// TIA Portal V19 export
FUNCTION_BLOCK "RUA_R4"   // FB22, LAD
{ S7_Optimized_Access := 'TRUE' }
// stored: MemoryReserve 100, SetENOAutomatically false
   VAR
      START_Instance { S7_SetPoint := 'True'} : "START";
      "HEAT/COOL_Instance" { S7_SetPoint := 'True'} : "HEAT/COOL";
      "AUTO_COOLING_UTIITY SELECTION_Instance" { S7_SetPoint := 'True'} : "AUTO_COOLING_UTIITY SELECTION";
      AUTO_HEATING_SELECTION_Instance { S7_SetPoint := 'True'} : "AUTO_HEATING_SELECTION";
      "SEMI/_AUTO_Instance" { S7_SetPoint := 'True'} : "SEMI/_AUTO";
      COOLING_PROCESS_Instance { S7_SetPoint := 'True'} : "COOLING_PROCESS";
      HEATING_PROCEES_Instance { S7_SetPoint := 'True'} : "HEATING_PROCEES";
      RAMP_Instance { S7_SetPoint := 'True'} : "RAMP";
   END_VAR
BEGIN

REGION Network 1: START
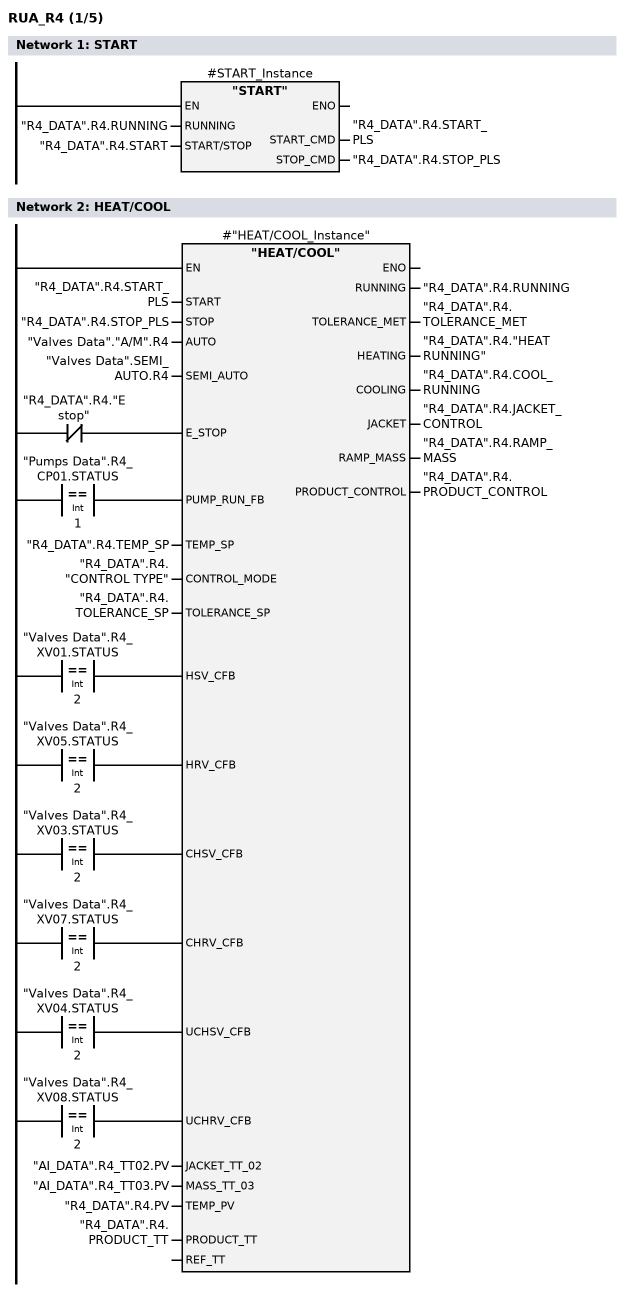
   RUNG wire#powerrail
      #START_Instance(RUNNING := "R4_DATA".R4.RUNNING, "START/STOP" := "R4_DATA".R4.START, START_CMD => "R4_DATA".R4.START_PLS, STOP_CMD => "R4_DATA".R4.STOP_PLS)
   END_RUNG
   // the same network as SCL:
   #START_Instance(RUNNING := "R4_DATA".R4.RUNNING,   // "START"
                   "START/STOP" := "R4_DATA".R4.START,
                   START_CMD => "R4_DATA".R4.START_PLS,
                   STOP_CMD => "R4_DATA".R4.STOP_PLS);
END_REGION

REGION Network 2: HEAT/COOL
   RUNG wire#powerrail
      #"HEAT/COOL_Instance"(E_STOP := wire#w1, PUMP_RUN_FB := wire#w2, HSV_CFB := wire#w3, HRV_CFB := wire#w4, CHSV_CFB := wire#w5, CHRV_CFB := wire#w6, UCHSV_CFB := wire#w7, UCHRV_CFB := wire#w8, START := "R4_DATA".R4.START_PLS, STOP := "R4_DATA".R4.STOP_PLS, AUTO := "Valves Data"."A/M".R4, SEMI_AUTO := "Valves Data".SEMI_AUTO.R4, TEMP_SP := "R4_DATA".R4.TEMP_SP, CONTROL_MODE := "R4_DATA".R4."CONTROL TYPE", TOLERANCE_SP := "R4_DATA".R4.TOLERANCE_SP, JACKET_TT_02 := "AI_DATA".R4_TT02.PV, MASS_TT_03 := "AI_DATA".R4_TT03.PV, TEMP_PV := "R4_DATA".R4.PV, PRODUCT_TT := "R4_DATA".R4.PRODUCT_TT, REF_TT :=, RUNNING => "R4_DATA".R4.RUNNING, TOLERANCE_MET => "R4_DATA".R4.TOLERANCE_MET, HEATING => "R4_DATA".R4."HEAT RUNNING", COOLING => "R4_DATA".R4.COOL_RUNNING, JACKET => "R4_DATA".R4.JACKET_CONTROL, RAMP_MASS => "R4_DATA".R4.RAMP_MASS, PRODUCT_CONTROL => "R4_DATA".R4.PRODUCT_CONTROL)
   END_RUNG
   RUNG wire#powerrail
      I_Contact( "R4_DATA".R4."E stop" )
   END_RUNG wire#w1
   RUNG wire#powerrail
      { S7_Templates := "SrcType := Int" } EQ_Contact(in1 := "Pumps Data".R4_CP01.STATUS, in2 := 1)
   END_RUNG wire#w2
   RUNG wire#powerrail
      { S7_Templates := "SrcType := Int" } EQ_Contact(in1 := "Valves Data".R4_XV01.STATUS, in2 := 2)
   END_RUNG wire#w3
   RUNG wire#powerrail
      { S7_Templates := "SrcType := Int" } EQ_Contact(in1 := "Valves Data".R4_XV05.STATUS, in2 := 2)
   END_RUNG wire#w4
   RUNG wire#powerrail
      { S7_Templates := "SrcType := Int" } EQ_Contact(in1 := "Valves Data".R4_XV03.STATUS, in2 := 2)
   END_RUNG wire#w5
   RUNG wire#powerrail
      { S7_Templates := "SrcType := Int" } EQ_Contact(in1 := "Valves Data".R4_XV07.STATUS, in2 := 2)
   END_RUNG wire#w6
   RUNG wire#powerrail
      { S7_Templates := "SrcType := Int" } EQ_Contact(in1 := "Valves Data".R4_XV04.STATUS, in2 := 2)
   END_RUNG wire#w7
   RUNG wire#powerrail
      { S7_Templates := "SrcType := Int" } EQ_Contact(in1 := "Valves Data".R4_XV08.STATUS, in2 := 2)
   END_RUNG wire#w8
   // the same network as SCL:
   #"HEAT/COOL_Instance"(START := "R4_DATA".R4.START_PLS,   // "HEAT/COOL"
                         STOP := "R4_DATA".R4.STOP_PLS,
                         AUTO := "Valves Data"."A/M".R4,
                         SEMI_AUTO := "Valves Data".SEMI_AUTO.R4,
                         E_STOP := NOT "R4_DATA".R4."E stop",
                         PUMP_RUN_FB := "Pumps Data".R4_CP01.STATUS = 1,
                         TEMP_SP := "R4_DATA".R4.TEMP_SP,
                         CONTROL_MODE := "R4_DATA".R4."CONTROL TYPE",
                         TOLERANCE_SP := "R4_DATA".R4.TOLERANCE_SP,
                         HSV_CFB := "Valves Data".R4_XV01.STATUS = 2,
                         HRV_CFB := "Valves Data".R4_XV05.STATUS = 2,
                         CHSV_CFB := "Valves Data".R4_XV03.STATUS = 2,
                         CHRV_CFB := "Valves Data".R4_XV07.STATUS = 2,
                         UCHSV_CFB := "Valves Data".R4_XV04.STATUS = 2,
                         UCHRV_CFB := "Valves Data".R4_XV08.STATUS = 2,
                         JACKET_TT_02 := "AI_DATA".R4_TT02.PV,
                         MASS_TT_03 := "AI_DATA".R4_TT03.PV,
                         TEMP_PV := "R4_DATA".R4.PV,
                         PRODUCT_TT := "R4_DATA".R4.PRODUCT_TT,
                         RUNNING => "R4_DATA".R4.RUNNING,
                         TOLERANCE_MET => "R4_DATA".R4.TOLERANCE_MET,
                         HEATING => "R4_DATA".R4."HEAT RUNNING",
                         COOLING => "R4_DATA".R4.COOL_RUNNING,
                         JACKET => "R4_DATA".R4.JACKET_CONTROL,
                         RAMP_MASS => "R4_DATA".R4.RAMP_MASS,
                         PRODUCT_CONTROL => "R4_DATA".R4.PRODUCT_CONTROL);
END_REGION

REGION Network 3: AUTO_COOLING
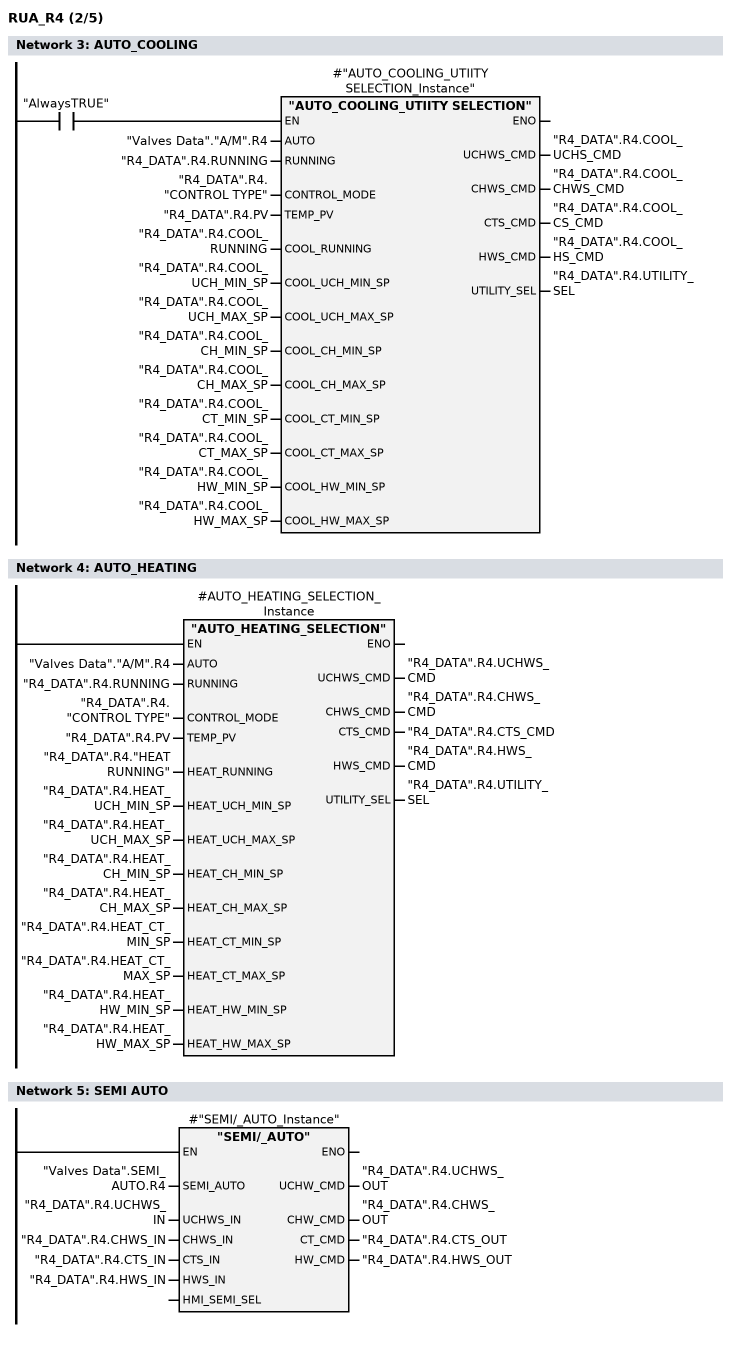
   RUNG wire#powerrail
      Contact( "AlwaysTRUE" )
      #"AUTO_COOLING_UTIITY SELECTION_Instance"(AUTO := "Valves Data"."A/M".R4, RUNNING := "R4_DATA".R4.RUNNING, CONTROL_MODE := "R4_DATA".R4."CONTROL TYPE", TEMP_PV := "R4_DATA".R4.PV, COOL_RUNNING := "R4_DATA".R4.COOL_RUNNING, COOL_UCH_MIN_SP := "R4_DATA".R4.COOL_UCH_MIN_SP, COOL_UCH_MAX_SP := "R4_DATA".R4.COOL_UCH_MAX_SP, COOL_CH_MIN_SP := "R4_DATA".R4.COOL_CH_MIN_SP, COOL_CH_MAX_SP := "R4_DATA".R4.COOL_CH_MAX_SP, COOL_CT_MIN_SP := "R4_DATA".R4.COOL_CT_MIN_SP, COOL_CT_MAX_SP := "R4_DATA".R4.COOL_CT_MAX_SP, COOL_HW_MIN_SP := "R4_DATA".R4.COOL_HW_MIN_SP, COOL_HW_MAX_SP := "R4_DATA".R4.COOL_HW_MAX_SP, UCHWS_CMD => "R4_DATA".R4.COOL_UCHS_CMD, CHWS_CMD => "R4_DATA".R4.COOL_CHWS_CMD, CTS_CMD => "R4_DATA".R4.COOL_CS_CMD, HWS_CMD => "R4_DATA".R4.COOL_HS_CMD, UTILITY_SEL => "R4_DATA".R4.UTILITY_SEL)
   END_RUNG
   // the same network as SCL:
   IF "AlwaysTRUE" THEN
       #"AUTO_COOLING_UTIITY SELECTION_Instance"(AUTO := "Valves Data"."A/M".R4,   // "AUTO_COOLING_UTIITY SELECTION"
                               RUNNING := "R4_DATA".R4.RUNNING,
                               CONTROL_MODE := "R4_DATA".R4."CONTROL TYPE",
                               TEMP_PV := "R4_DATA".R4.PV,
                               COOL_RUNNING := "R4_DATA".R4.COOL_RUNNING,
                               COOL_UCH_MIN_SP := "R4_DATA".R4.COOL_UCH_MIN_SP,
                               COOL_UCH_MAX_SP := "R4_DATA".R4.COOL_UCH_MAX_SP,
                               COOL_CH_MIN_SP := "R4_DATA".R4.COOL_CH_MIN_SP,
                               COOL_CH_MAX_SP := "R4_DATA".R4.COOL_CH_MAX_SP,
                               COOL_CT_MIN_SP := "R4_DATA".R4.COOL_CT_MIN_SP,
                               COOL_CT_MAX_SP := "R4_DATA".R4.COOL_CT_MAX_SP,
                               COOL_HW_MIN_SP := "R4_DATA".R4.COOL_HW_MIN_SP,
                               COOL_HW_MAX_SP := "R4_DATA".R4.COOL_HW_MAX_SP,
                               UCHWS_CMD => "R4_DATA".R4.COOL_UCHS_CMD,
                               CHWS_CMD => "R4_DATA".R4.COOL_CHWS_CMD,
                               CTS_CMD => "R4_DATA".R4.COOL_CS_CMD,
                               HWS_CMD => "R4_DATA".R4.COOL_HS_CMD,
                               UTILITY_SEL => "R4_DATA".R4.UTILITY_SEL);
   END_IF;
END_REGION

REGION Network 4: AUTO_HEATING
   RUNG wire#powerrail
      #AUTO_HEATING_SELECTION_Instance(AUTO := "Valves Data"."A/M".R4, RUNNING := "R4_DATA".R4.RUNNING, CONTROL_MODE := "R4_DATA".R4."CONTROL TYPE", TEMP_PV := "R4_DATA".R4.PV, HEAT_RUNNING := "R4_DATA".R4."HEAT RUNNING", HEAT_UCH_MIN_SP := "R4_DATA".R4.HEAT_UCH_MIN_SP, HEAT_UCH_MAX_SP := "R4_DATA".R4.HEAT_UCH_MAX_SP, HEAT_CH_MIN_SP := "R4_DATA".R4.HEAT_CH_MIN_SP, HEAT_CH_MAX_SP := "R4_DATA".R4.HEAT_CH_MAX_SP, HEAT_CT_MIN_SP := "R4_DATA".R4.HEAT_CT_MIN_SP, HEAT_CT_MAX_SP := "R4_DATA".R4.HEAT_CT_MAX_SP, HEAT_HW_MIN_SP := "R4_DATA".R4.HEAT_HW_MIN_SP, HEAT_HW_MAX_SP := "R4_DATA".R4.HEAT_HW_MAX_SP, UCHWS_CMD => "R4_DATA".R4.UCHWS_CMD, CHWS_CMD => "R4_DATA".R4.CHWS_CMD, CTS_CMD => "R4_DATA".R4.CTS_CMD, HWS_CMD => "R4_DATA".R4.HWS_CMD, UTILITY_SEL => "R4_DATA".R4.UTILITY_SEL)
   END_RUNG
   // the same network as SCL:
   #AUTO_HEATING_SELECTION_Instance(AUTO := "Valves Data"."A/M".R4,   // "AUTO_HEATING_SELECTION"
                           RUNNING := "R4_DATA".R4.RUNNING,
                           CONTROL_MODE := "R4_DATA".R4."CONTROL TYPE",
                           TEMP_PV := "R4_DATA".R4.PV,
                           HEAT_RUNNING := "R4_DATA".R4."HEAT RUNNING",
                           HEAT_UCH_MIN_SP := "R4_DATA".R4.HEAT_UCH_MIN_SP,
                           HEAT_UCH_MAX_SP := "R4_DATA".R4.HEAT_UCH_MAX_SP,
                           HEAT_CH_MIN_SP := "R4_DATA".R4.HEAT_CH_MIN_SP,
                           HEAT_CH_MAX_SP := "R4_DATA".R4.HEAT_CH_MAX_SP,
                           HEAT_CT_MIN_SP := "R4_DATA".R4.HEAT_CT_MIN_SP,
                           HEAT_CT_MAX_SP := "R4_DATA".R4.HEAT_CT_MAX_SP,
                           HEAT_HW_MIN_SP := "R4_DATA".R4.HEAT_HW_MIN_SP,
                           HEAT_HW_MAX_SP := "R4_DATA".R4.HEAT_HW_MAX_SP,
                           UCHWS_CMD => "R4_DATA".R4.UCHWS_CMD,
                           CHWS_CMD => "R4_DATA".R4.CHWS_CMD,
                           CTS_CMD => "R4_DATA".R4.CTS_CMD,
                           HWS_CMD => "R4_DATA".R4.HWS_CMD,
                           UTILITY_SEL => "R4_DATA".R4.UTILITY_SEL);
END_REGION

REGION Network 5: SEMI AUTO
   RUNG wire#powerrail
      #"SEMI/_AUTO_Instance"(SEMI_AUTO := "Valves Data".SEMI_AUTO.R4, UCHWS_IN := "R4_DATA".R4.UCHWS_IN, CHWS_IN := "R4_DATA".R4.CHWS_IN, CTS_IN := "R4_DATA".R4.CTS_IN, HWS_IN := "R4_DATA".R4.HWS_IN, UCHW_CMD => "R4_DATA".R4.UCHWS_OUT, CHW_CMD => "R4_DATA".R4.CHWS_OUT, CT_CMD => "R4_DATA".R4.CTS_OUT, HW_CMD => "R4_DATA".R4.HWS_OUT, HMI_SEMI_SEL :=)
   END_RUNG
   // the same network as SCL:
   #"SEMI/_AUTO_Instance"(SEMI_AUTO := "Valves Data".SEMI_AUTO.R4,   // "SEMI/_AUTO"
                          UCHWS_IN := "R4_DATA".R4.UCHWS_IN,
                          CHWS_IN := "R4_DATA".R4.CHWS_IN,
                          CTS_IN := "R4_DATA".R4.CTS_IN,
                          HWS_IN := "R4_DATA".R4.HWS_IN,
                          UCHW_CMD => "R4_DATA".R4.UCHWS_OUT,
                          CHW_CMD => "R4_DATA".R4.CHWS_OUT,
                          CT_CMD => "R4_DATA".R4.CTS_OUT,
                          HW_CMD => "R4_DATA".R4.HWS_OUT);
END_REGION

REGION Network 6: COOLING_PROCESS
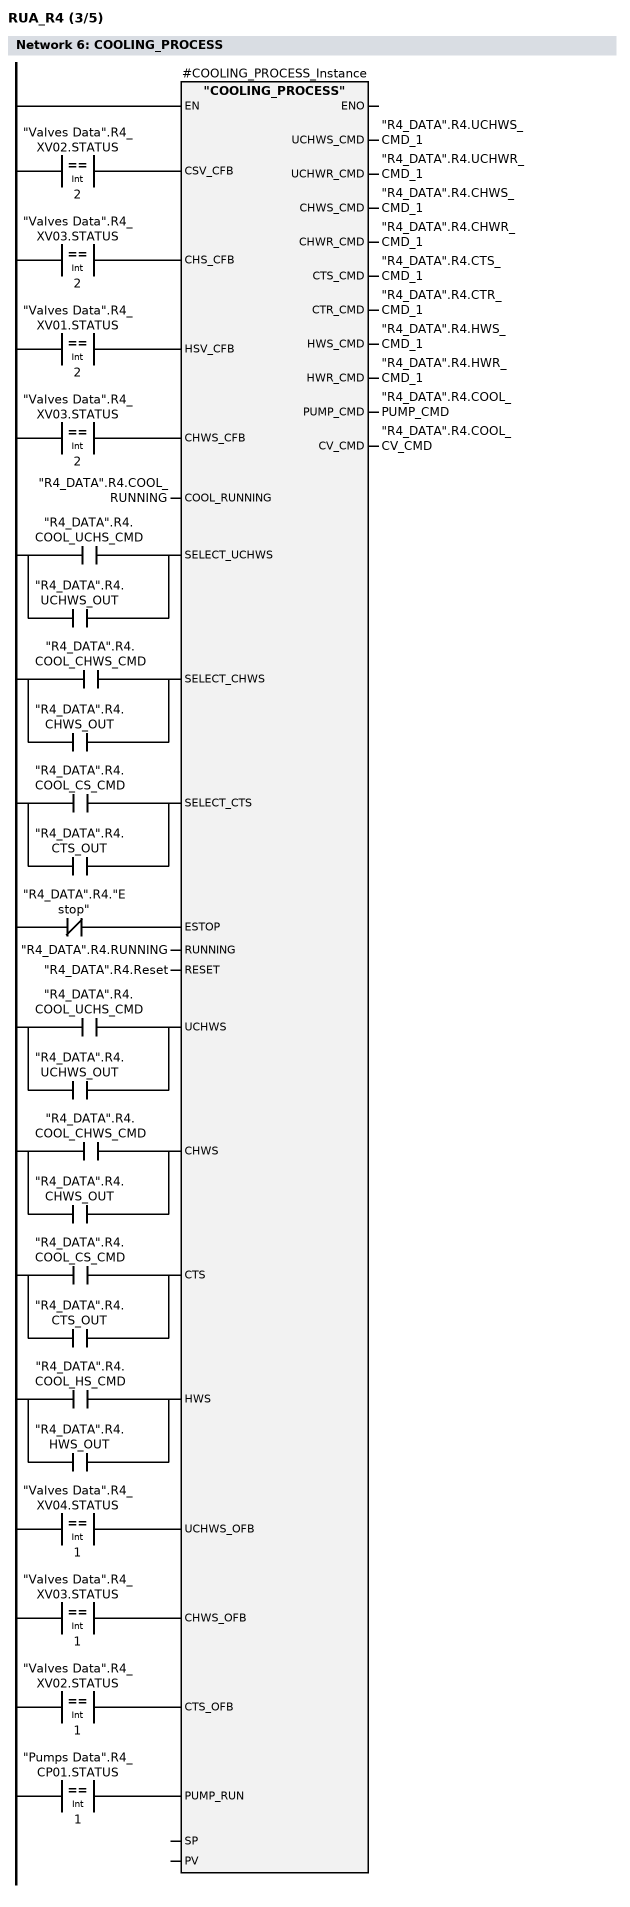
   RUNG wire#powerrail
      #COOLING_PROCESS_Instance(CSV_CFB := wire#w1, CHS_CFB := wire#w2, HSV_CFB := wire#w3, CHWS_CFB := wire#w4, SELECT_UCHWS := wire#w5, SELECT_CHWS := wire#w6, SELECT_CTS := wire#w7, ESTOP := wire#w8, UCHWS := wire#w9, CHWS := wire#w10, CTS := wire#w11, HWS := wire#w12, UCHWS_OFB := wire#w13, CHWS_OFB := wire#w14, CTS_OFB := wire#w15, PUMP_RUN := wire#w16, COOL_RUNNING := "R4_DATA".R4.COOL_RUNNING, RUNNING := "R4_DATA".R4.RUNNING, RESET := "R4_DATA".R4.Reset, SP :=, PV :=, UCHWS_CMD => "R4_DATA".R4.UCHWS_CMD_1, UCHWR_CMD => "R4_DATA".R4.UCHWR_CMD_1, CHWS_CMD => "R4_DATA".R4.CHWS_CMD_1, CHWR_CMD => "R4_DATA".R4.CHWR_CMD_1, CTS_CMD => "R4_DATA".R4.CTS_CMD_1, CTR_CMD => "R4_DATA".R4.CTR_CMD_1, HWS_CMD => "R4_DATA".R4.HWS_CMD_1, HWR_CMD => "R4_DATA".R4.HWR_CMD_1, PUMP_CMD => "R4_DATA".R4.COOL_PUMP_CMD, CV_CMD => "R4_DATA".R4.COOL_CV_CMD)
   END_RUNG
   RUNG wire#powerrail
      { S7_Templates := "SrcType := Int" } EQ_Contact(in1 := "Valves Data".R4_XV02.STATUS, in2 := 2)
   END_RUNG wire#w1
   RUNG wire#powerrail
      { S7_Templates := "SrcType := Int" } EQ_Contact(in1 := "Valves Data".R4_XV03.STATUS, in2 := 2)
   END_RUNG wire#w2
   RUNG wire#powerrail
      { S7_Templates := "SrcType := Int" } EQ_Contact(in1 := "Valves Data".R4_XV01.STATUS, in2 := 2)
   END_RUNG wire#w3
   RUNG wire#powerrail
      { S7_Templates := "SrcType := Int" } EQ_Contact(in1 := "Valves Data".R4_XV03.STATUS, in2 := 2)
   END_RUNG wire#w4
   RUNG wire#powerrail
      Contact( "R4_DATA".R4.COOL_UCHS_CMD )
   END_RUNG wire#w5
   RUNG wire#powerrail
      Contact( "R4_DATA".R4.UCHWS_OUT )
   END_RUNG wire#w5
   RUNG wire#powerrail
      Contact( "R4_DATA".R4.COOL_CHWS_CMD )
   END_RUNG wire#w6
   RUNG wire#powerrail
      Contact( "R4_DATA".R4.CHWS_OUT )
   END_RUNG wire#w6
   RUNG wire#powerrail
      Contact( "R4_DATA".R4.COOL_CS_CMD )
   END_RUNG wire#w7
   RUNG wire#powerrail
      Contact( "R4_DATA".R4.CTS_OUT )
   END_RUNG wire#w7
   RUNG wire#powerrail
      I_Contact( "R4_DATA".R4."E stop" )
   END_RUNG wire#w8
   RUNG wire#powerrail
      Contact( "R4_DATA".R4.COOL_UCHS_CMD )
   END_RUNG wire#w9
   RUNG wire#powerrail
      Contact( "R4_DATA".R4.UCHWS_OUT )
   END_RUNG wire#w9
   RUNG wire#powerrail
      Contact( "R4_DATA".R4.COOL_CHWS_CMD )
   END_RUNG wire#w10
   RUNG wire#powerrail
      Contact( "R4_DATA".R4.CHWS_OUT )
   END_RUNG wire#w10
   RUNG wire#powerrail
      Contact( "R4_DATA".R4.COOL_CS_CMD )
   END_RUNG wire#w11
   RUNG wire#powerrail
      Contact( "R4_DATA".R4.CTS_OUT )
   END_RUNG wire#w11
   RUNG wire#powerrail
      Contact( "R4_DATA".R4.COOL_HS_CMD )
   END_RUNG wire#w12
   RUNG wire#powerrail
      Contact( "R4_DATA".R4.HWS_OUT )
   END_RUNG wire#w12
   RUNG wire#powerrail
      { S7_Templates := "SrcType := Int" } EQ_Contact(in1 := "Valves Data".R4_XV04.STATUS, in2 := 1)
   END_RUNG wire#w13
   RUNG wire#powerrail
      { S7_Templates := "SrcType := Int" } EQ_Contact(in1 := "Valves Data".R4_XV03.STATUS, in2 := 1)
   END_RUNG wire#w14
   RUNG wire#powerrail
      { S7_Templates := "SrcType := Int" } EQ_Contact(in1 := "Valves Data".R4_XV02.STATUS, in2 := 1)
   END_RUNG wire#w15
   RUNG wire#powerrail
      { S7_Templates := "SrcType := Int" } EQ_Contact(in1 := "Pumps Data".R4_CP01.STATUS, in2 := 1)
   END_RUNG wire#w16
   // the same network as SCL:
   #COOLING_PROCESS_Instance(CSV_CFB := "Valves Data".R4_XV02.STATUS = 2,   // "COOLING_PROCESS"
                           CHS_CFB := "Valves Data".R4_XV03.STATUS = 2,
                           HSV_CFB := "Valves Data".R4_XV01.STATUS = 2,
                           CHWS_CFB := "Valves Data".R4_XV03.STATUS = 2,
                           COOL_RUNNING := "R4_DATA".R4.COOL_RUNNING,
                           SELECT_UCHWS := "R4_DATA".R4.COOL_UCHS_CMD OR "R4_DATA".R4.UCHWS_OUT,
                           SELECT_CHWS := "R4_DATA".R4.COOL_CHWS_CMD OR "R4_DATA".R4.CHWS_OUT,
                           SELECT_CTS := "R4_DATA".R4.COOL_CS_CMD OR "R4_DATA".R4.CTS_OUT,
                           ESTOP := NOT "R4_DATA".R4."E stop",
                           RUNNING := "R4_DATA".R4.RUNNING,
                           RESET := "R4_DATA".R4.Reset,
                           UCHWS := "R4_DATA".R4.COOL_UCHS_CMD OR "R4_DATA".R4.UCHWS_OUT,
                           CHWS := "R4_DATA".R4.COOL_CHWS_CMD OR "R4_DATA".R4.CHWS_OUT,
                           CTS := "R4_DATA".R4.COOL_CS_CMD OR "R4_DATA".R4.CTS_OUT,
                           HWS := "R4_DATA".R4.COOL_HS_CMD OR "R4_DATA".R4.HWS_OUT,
                           UCHWS_OFB := "Valves Data".R4_XV04.STATUS = 1,
                           CHWS_OFB := "Valves Data".R4_XV03.STATUS = 1,
                           CTS_OFB := "Valves Data".R4_XV02.STATUS = 1,
                           PUMP_RUN := "Pumps Data".R4_CP01.STATUS = 1,
                           UCHWS_CMD => "R4_DATA".R4.UCHWS_CMD_1,
                           UCHWR_CMD => "R4_DATA".R4.UCHWR_CMD_1,
                           CHWS_CMD => "R4_DATA".R4.CHWS_CMD_1,
                           CHWR_CMD => "R4_DATA".R4.CHWR_CMD_1,
                           CTS_CMD => "R4_DATA".R4.CTS_CMD_1,
                           CTR_CMD => "R4_DATA".R4.CTR_CMD_1,
                           HWS_CMD => "R4_DATA".R4.HWS_CMD_1,
                           HWR_CMD => "R4_DATA".R4.HWR_CMD_1,
                           PUMP_CMD => "R4_DATA".R4.COOL_PUMP_CMD,
                           CV_CMD => "R4_DATA".R4.COOL_CV_CMD);
END_REGION

REGION Network 7: HEATING PROCESS
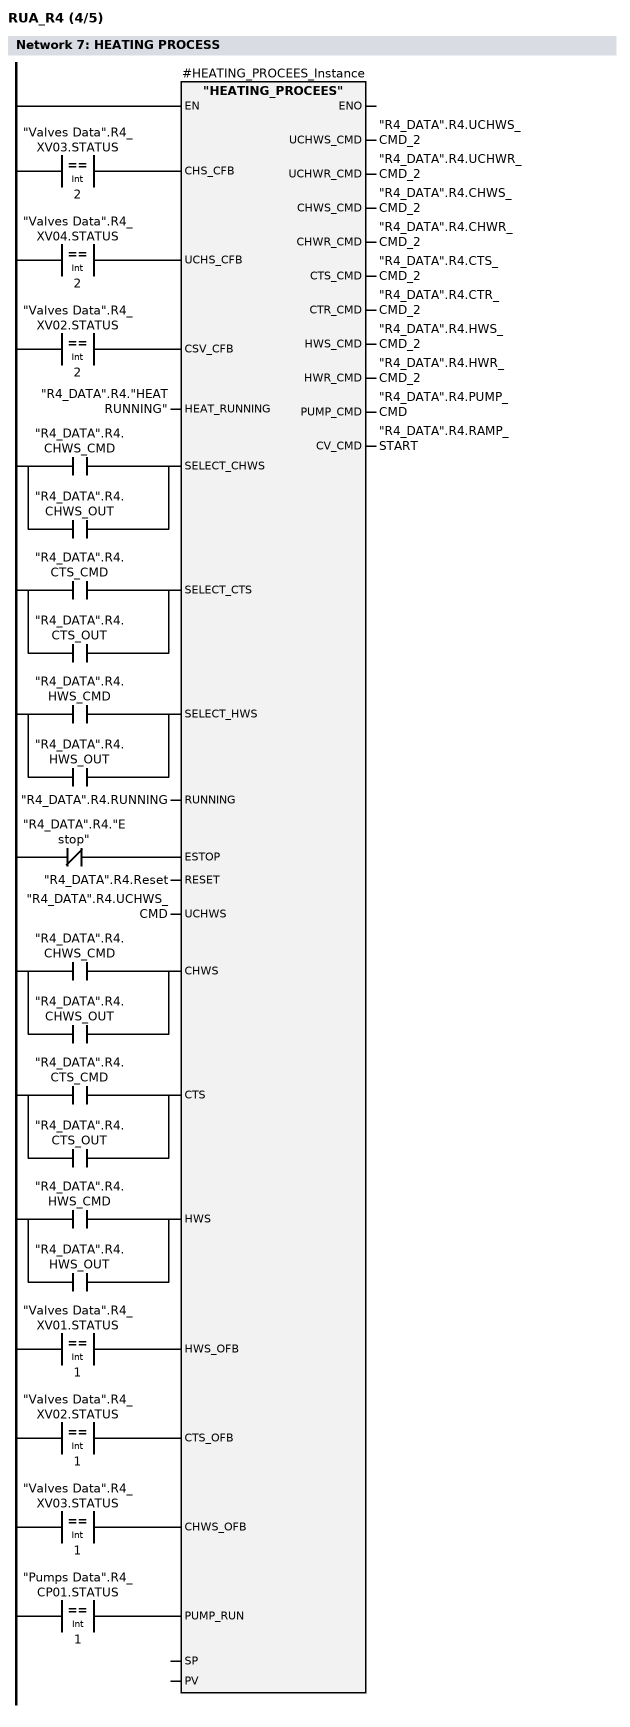
   RUNG wire#powerrail
      #HEATING_PROCEES_Instance(CHS_CFB := wire#w1, UCHS_CFB := wire#w2, CSV_CFB := wire#w3, SELECT_CHWS := wire#w4, SELECT_CTS := wire#w5, SELECT_HWS := wire#w6, ESTOP := wire#w7, CHWS := wire#w8, CTS := wire#w9, HWS := wire#w10, HWS_OFB := wire#w11, CTS_OFB := wire#w12, CHWS_OFB := wire#w13, PUMP_RUN := wire#w14, HEAT_RUNNING := "R4_DATA".R4."HEAT RUNNING", RUNNING := "R4_DATA".R4.RUNNING, RESET := "R4_DATA".R4.Reset, UCHWS := "R4_DATA".R4.UCHWS_CMD, SP :=, PV :=, UCHWS_CMD => "R4_DATA".R4.UCHWS_CMD_2, UCHWR_CMD => "R4_DATA".R4.UCHWR_CMD_2, CHWS_CMD => "R4_DATA".R4.CHWS_CMD_2, CHWR_CMD => "R4_DATA".R4.CHWR_CMD_2, CTS_CMD => "R4_DATA".R4.CTS_CMD_2, CTR_CMD => "R4_DATA".R4.CTR_CMD_2, HWS_CMD => "R4_DATA".R4.HWS_CMD_2, HWR_CMD => "R4_DATA".R4.HWR_CMD_2, PUMP_CMD => "R4_DATA".R4.PUMP_CMD, CV_CMD => "R4_DATA".R4.RAMP_START)
   END_RUNG
   RUNG wire#powerrail
      { S7_Templates := "SrcType := Int" } EQ_Contact(in1 := "Valves Data".R4_XV03.STATUS, in2 := 2)
   END_RUNG wire#w1
   RUNG wire#powerrail
      { S7_Templates := "SrcType := Int" } EQ_Contact(in1 := "Valves Data".R4_XV04.STATUS, in2 := 2)
   END_RUNG wire#w2
   RUNG wire#powerrail
      { S7_Templates := "SrcType := Int" } EQ_Contact(in1 := "Valves Data".R4_XV02.STATUS, in2 := 2)
   END_RUNG wire#w3
   RUNG wire#powerrail
      Contact( "R4_DATA".R4.CHWS_CMD )
   END_RUNG wire#w4
   RUNG wire#powerrail
      Contact( "R4_DATA".R4.CHWS_OUT )
   END_RUNG wire#w4
   RUNG wire#powerrail
      Contact( "R4_DATA".R4.CTS_CMD )
   END_RUNG wire#w5
   RUNG wire#powerrail
      Contact( "R4_DATA".R4.CTS_OUT )
   END_RUNG wire#w5
   RUNG wire#powerrail
      Contact( "R4_DATA".R4.HWS_CMD )
   END_RUNG wire#w6
   RUNG wire#powerrail
      Contact( "R4_DATA".R4.HWS_OUT )
   END_RUNG wire#w6
   RUNG wire#powerrail
      I_Contact( "R4_DATA".R4."E stop" )
   END_RUNG wire#w7
   RUNG wire#powerrail
      Contact( "R4_DATA".R4.CHWS_CMD )
   END_RUNG wire#w8
   RUNG wire#powerrail
      Contact( "R4_DATA".R4.CHWS_OUT )
   END_RUNG wire#w8
   RUNG wire#powerrail
      Contact( "R4_DATA".R4.CTS_CMD )
   END_RUNG wire#w9
   RUNG wire#powerrail
      Contact( "R4_DATA".R4.CTS_OUT )
   END_RUNG wire#w9
   RUNG wire#powerrail
      Contact( "R4_DATA".R4.HWS_CMD )
   END_RUNG wire#w10
   RUNG wire#powerrail
      Contact( "R4_DATA".R4.HWS_OUT )
   END_RUNG wire#w10
   RUNG wire#powerrail
      { S7_Templates := "SrcType := Int" } EQ_Contact(in1 := "Valves Data".R4_XV01.STATUS, in2 := 1)
   END_RUNG wire#w11
   RUNG wire#powerrail
      { S7_Templates := "SrcType := Int" } EQ_Contact(in1 := "Valves Data".R4_XV02.STATUS, in2 := 1)
   END_RUNG wire#w12
   RUNG wire#powerrail
      { S7_Templates := "SrcType := Int" } EQ_Contact(in1 := "Valves Data".R4_XV03.STATUS, in2 := 1)
   END_RUNG wire#w13
   RUNG wire#powerrail
      { S7_Templates := "SrcType := Int" } EQ_Contact(in1 := "Pumps Data".R4_CP01.STATUS, in2 := 1)
   END_RUNG wire#w14
   // the same network as SCL:
   #HEATING_PROCEES_Instance(CHS_CFB := "Valves Data".R4_XV03.STATUS = 2,   // "HEATING_PROCEES"
                           UCHS_CFB := "Valves Data".R4_XV04.STATUS = 2,
                           CSV_CFB := "Valves Data".R4_XV02.STATUS = 2,
                           HEAT_RUNNING := "R4_DATA".R4."HEAT RUNNING",
                           SELECT_CHWS := "R4_DATA".R4.CHWS_CMD OR "R4_DATA".R4.CHWS_OUT,
                           SELECT_CTS := "R4_DATA".R4.CTS_CMD OR "R4_DATA".R4.CTS_OUT,
                           SELECT_HWS := "R4_DATA".R4.HWS_CMD OR "R4_DATA".R4.HWS_OUT,
                           RUNNING := "R4_DATA".R4.RUNNING,
                           ESTOP := NOT "R4_DATA".R4."E stop",
                           RESET := "R4_DATA".R4.Reset,
                           UCHWS := "R4_DATA".R4.UCHWS_CMD,
                           CHWS := "R4_DATA".R4.CHWS_CMD OR "R4_DATA".R4.CHWS_OUT,
                           CTS := "R4_DATA".R4.CTS_CMD OR "R4_DATA".R4.CTS_OUT,
                           HWS := "R4_DATA".R4.HWS_CMD OR "R4_DATA".R4.HWS_OUT,
                           HWS_OFB := "Valves Data".R4_XV01.STATUS = 1,
                           CTS_OFB := "Valves Data".R4_XV02.STATUS = 1,
                           CHWS_OFB := "Valves Data".R4_XV03.STATUS = 1,
                           PUMP_RUN := "Pumps Data".R4_CP01.STATUS = 1,
                           UCHWS_CMD => "R4_DATA".R4.UCHWS_CMD_2,
                           UCHWR_CMD => "R4_DATA".R4.UCHWR_CMD_2,
                           CHWS_CMD => "R4_DATA".R4.CHWS_CMD_2,
                           CHWR_CMD => "R4_DATA".R4.CHWR_CMD_2,
                           CTS_CMD => "R4_DATA".R4.CTS_CMD_2,
                           CTR_CMD => "R4_DATA".R4.CTR_CMD_2,
                           HWS_CMD => "R4_DATA".R4.HWS_CMD_2,
                           HWR_CMD => "R4_DATA".R4.HWR_CMD_2,
                           PUMP_CMD => "R4_DATA".R4.PUMP_CMD,
                           CV_CMD => "R4_DATA".R4.RAMP_START);
END_REGION

REGION Network 8: RAMP
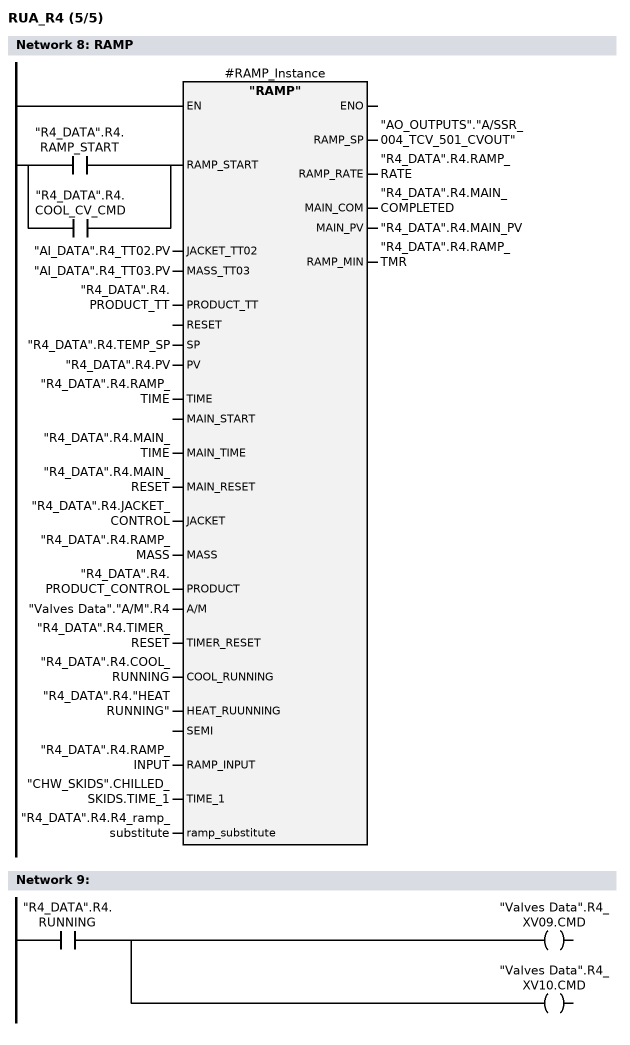
   RUNG wire#powerrail
      #RAMP_Instance(RAMP_START := wire#w1, JACKET_TT02 := "AI_DATA".R4_TT02.PV, MASS_TT03 := "AI_DATA".R4_TT03.PV, PRODUCT_TT := "R4_DATA".R4.PRODUCT_TT, RESET :=, SP := "R4_DATA".R4.TEMP_SP, PV := "R4_DATA".R4.PV, "TIME" := "R4_DATA".R4.RAMP_TIME, MAIN_START :=, MAIN_TIME := "R4_DATA".R4.MAIN_TIME, MAIN_RESET := "R4_DATA".R4.MAIN_RESET, JACKET := "R4_DATA".R4.JACKET_CONTROL, MASS := "R4_DATA".R4.RAMP_MASS, PRODUCT := "R4_DATA".R4.PRODUCT_CONTROL, "A/M" := "Valves Data"."A/M".R4, TIMER_RESET := "R4_DATA".R4.TIMER_RESET, COOL_RUNNING := "R4_DATA".R4.COOL_RUNNING, HEAT_RUUNNING := "R4_DATA".R4."HEAT RUNNING", RAMP_INPUT := "R4_DATA".R4.RAMP_INPUT, TIME_1 := "CHW_SKIDS".CHILLED_SKIDS.TIME_1, ramp_substitute := "R4_DATA".R4.R4_ramp_substitute, RAMP_SP => "AO_OUTPUTS"."A/SSR_004_TCV_501_CVOUT", RAMP_RATE => "R4_DATA".R4.RAMP_RATE, MAIN_COM => "R4_DATA".R4.MAIN_COMPLETED, MAIN_PV => "R4_DATA".R4.MAIN_PV, RAMP_MIN => "R4_DATA".R4.RAMP_TMR, SEMI :=)
   END_RUNG
   RUNG wire#powerrail
      Contact( "R4_DATA".R4.RAMP_START )
   END_RUNG wire#w1
   RUNG wire#powerrail
      Contact( "R4_DATA".R4.COOL_CV_CMD )
   END_RUNG wire#w1
   // the same network as SCL:
   #RAMP_Instance(RAMP_START := "R4_DATA".R4.RAMP_START OR "R4_DATA".R4.COOL_CV_CMD,   // "RAMP"
                  JACKET_TT02 := "AI_DATA".R4_TT02.PV,
                  MASS_TT03 := "AI_DATA".R4_TT03.PV,
                  PRODUCT_TT := "R4_DATA".R4.PRODUCT_TT,
                  SP := "R4_DATA".R4.TEMP_SP,
                  PV := "R4_DATA".R4.PV,
                  "TIME" := "R4_DATA".R4.RAMP_TIME,
                  MAIN_TIME := "R4_DATA".R4.MAIN_TIME,
                  MAIN_RESET := "R4_DATA".R4.MAIN_RESET,
                  JACKET := "R4_DATA".R4.JACKET_CONTROL,
                  MASS := "R4_DATA".R4.RAMP_MASS,
                  PRODUCT := "R4_DATA".R4.PRODUCT_CONTROL,
                  "A/M" := "Valves Data"."A/M".R4,
                  TIMER_RESET := "R4_DATA".R4.TIMER_RESET,
                  COOL_RUNNING := "R4_DATA".R4.COOL_RUNNING,
                  HEAT_RUUNNING := "R4_DATA".R4."HEAT RUNNING",
                  RAMP_INPUT := "R4_DATA".R4.RAMP_INPUT,
                  TIME_1 := "CHW_SKIDS".CHILLED_SKIDS.TIME_1,
                  ramp_substitute := "R4_DATA".R4.R4_ramp_substitute,
                  RAMP_SP => "AO_OUTPUTS"."A/SSR_004_TCV_501_CVOUT",
                  RAMP_RATE => "R4_DATA".R4.RAMP_RATE,
                  MAIN_COM => "R4_DATA".R4.MAIN_COMPLETED,
                  MAIN_PV => "R4_DATA".R4.MAIN_PV,
                  RAMP_MIN => "R4_DATA".R4.RAMP_TMR);
END_REGION

REGION Network 9
   RUNG wire#powerrail
      Contact( "R4_DATA".R4.RUNNING )
      wire#w1
      Coil( "Valves Data".R4_XV09.CMD )
   END_RUNG
   RUNG wire#w1
      Coil( "Valves Data".R4_XV10.CMD )
   END_RUNG
   // the same network as SCL:
   "Valves Data".R4_XV09.CMD := "R4_DATA".R4.RUNNING;
   "Valves Data".R4_XV10.CMD := "R4_DATA".R4.RUNNING;
END_REGION
END_FUNCTION_BLOCK
